// TIA Portal V21 export
// export: Created 2000-01-01T00:00:00.0000000Z, ExportSetting None
TYPE "UDT_HMI_FIO_TankLevelPID"
   STRUCT
      bManualMode { ExternalWritable := 'False'} : Bool;   // TRUE: 手动开度给定模式, FALSE: 自动PID闭环模式
      bResetCmd { ExternalWritable := 'False'} : Bool;   // HMI复位积分项与报警
      rSetpoint { ExternalWritable := 'False'} : Real;   // 液位设定值 SP (0.0..300.0 cm，默认 150.0)
      rKp { ExternalWritable := 'False'} : Real;   // 比例增益 Kp (默认 2.0)
      rKi { ExternalWritable := 'False'} : Real;   // 积分增益 Ki (1/s，默认 0.2)
      rKd { ExternalWritable := 'False'} : Real;   // 微分增益 Kd (s，默认 0.05)
      rDeadband { ExternalWritable := 'False'} : Real;   // 稳态误差死区 (cm，默认 0.5)
      rManualFillValve { ExternalWritable := 'False'} : Real;   // 手动进水阀开度给定 (0.0..10.0V)
      rManualDischargeValve { ExternalWritable := 'False'} : Real;   // 手动排水阀开度给定 (0.0..10.0V)
      rCurrentLevel { ExternalWritable := 'False'} : Real;   // 状态反馈：当前实际液位 PV (0.0..300.0 cm)
      rControlError { ExternalWritable := 'False'} : Real;   // 状态反馈：当前偏差 e = SP - PV
      rFillValveOut { ExternalWritable := 'False'} : Real;   // 状态反馈：进水比例阀输出电压 (0.0..10.0V)
      rDischargeValveOut { ExternalWritable := 'False'} : Real;   // 状态反馈：排水比例阀输出电压 (0.0..10.0V)
      bHighLevelAlarm { ExternalWritable := 'False'} : Bool;   // 状态反馈：高液位溢流联锁报警
      bLowLevelAlarm { ExternalWritable := 'False'} : Bool;   // 状态反馈：低液位干烧报警
      wStatus { ExternalWritable := 'False'} : Word;   // 状态码：16#0000正常, 16#7000停机, 16#8200采样周期非法, 16#8401高液位溢流保护, 16#8402急停切断
   END_STRUCT;
END_TYPE
